// Probe for MONETcommon#17: does a function block instance declared in a METHOD's plain VAR keep its state between
// calls? Each pair of methods is identical except for VAR versus VAR_INST (the control).
FUNCTION_BLOCK FB_MethodVarProbe
VAR
END_VAR

METHOD CountVar : INT
VAR
	n	: INT;
END_VAR
n := n + 1;
CountVar := n;
END_METHOD

METHOD CountInst : INT
VAR_INST
	n	: INT;
END_VAR
n := n + 1;
CountInst := n;
END_METHOD

METHOD EdgeVar : BOOL
VAR_INPUT
	bClk	: BOOL;
END_VAR
VAR
	rtrig	: R_TRIG;
END_VAR
rtrig(CLK := bClk);
EdgeVar := rtrig.Q;
END_METHOD

METHOD EdgeInst : BOOL
VAR_INPUT
	bClk	: BOOL;
END_VAR
VAR_INST
	rtrig	: R_TRIG;
END_VAR
rtrig(CLK := bClk);
EdgeInst := rtrig.Q;
END_METHOD

METHOD TimerVar : BOOL
VAR
	ton	: TON;
END_VAR
ton(IN := TRUE, PT := T#50MS);
TimerVar := ton.Q;
END_METHOD

METHOD TimerInst : BOOL
VAR_INST
	ton	: TON;
END_VAR
ton(IN := TRUE, PT := T#50MS);
TimerInst := ton.Q;
END_METHOD

END_FUNCTION_BLOCK

(* stored: Version 1.1.0.1, ProductVersion 3.1.4024.15
   POU FB_MethodVarProbe: Id {1e105a48-79a6-45e3-b089-6b8abaa15a00}, SpecialFunc None
   Method CountVar: Id {dc9e444b-8fa6-4c21-a6e4-74b8779c3418}
   Method CountInst: Id {f4542f34-7b6c-4e97-b05c-ffce4d996497}
   Method EdgeVar: Id {c5502fde-22b8-4b31-8ce5-17782a13ceb7}
   Method EdgeInst: Id {53cd8a8e-9935-4aa1-a2cf-073db6c2a02c}
   Method TimerVar: Id {12229898-2ab5-4a33-930f-e62e87b1b35d}
   Method TimerInst: Id {93179d1a-42a2-4033-8010-35a8bbf5a555} *)
